(* IEC 61131-3 sources: plcrex/tests/st_to_synchr_models, 21 files *)

(* ---- TC02.st ---- *)
FUNCTION_BLOCK TC02//_functionBlock
  VAR
    x0 : INT;
  END_VAR

  x0 := 0;
END_FUNCTION_BLOCK

(* ---- TC04.st ---- *)
FUNCTION_BLOCK TC04 //_inputs
  VAR_INPUT
    x0 : INT;
    x1 : INT := 6;
  END_VAR
  VAR
    x2 : INT;
  END_VAR

  x2 := x1;
END_FUNCTION_BLOCK

(* ---- TC05.st ---- *)
FUNCTION_BLOCK TC05 //_outputs
  VAR_OUTPUT
    y0 : INT;
    y1 : INT := 6;
  END_VAR
  VAR
    x2 : INT;
  END_VAR

  y0 := x2;
END_FUNCTION_BLOCK

(* ---- TC06.st ---- *)
FUNCTION_BLOCK TC06 //_in_outputs
  VAR_IN_OUT
    y0 : INT;
    y1 : INT;
  END_VAR

  y0 := y1;
END_FUNCTION_BLOCK

(* ---- TC07.st ---- *)
FUNCTION_BLOCK TC07 //_localVariables
  VAR
    x0 : INT;
    x1 : INT := 6;
  END_VAR

  x0 := x1;
END_FUNCTION_BLOCK

(* ---- TC08.st ---- *)
FUNCTION_BLOCK TC08 // _datatypes
  VAR
    x0 : BOOL;
    x1 : BOOL := TRUE;
    x2 : INT;
    x3 : INT := 2;
    x4 : REAL;
    x5 : REAL := 1.23;
    x7 : TIME;
    x8 : TIME := t#5s;
    x9 : ARRAY [1..2] OF BOOL;
    x10 : ARRAY [1..2] OF INT;
    x11 : ARRAY [1..2] OF REAL;
    x12 : ARRAY [1..2] OF TIME;
  END_VAR

  x0 := x1;
  x2 := x3;
  x4 := x5;
  x7 := x8;
  x9[0]:=TRUE;
  x10[0]:=2;
  x11[0]:=1.23;
  x12[0]:=t#2s;
END_FUNCTION_BLOCK

(* ---- TC09.st ---- *)
FUNCTION_BLOCK TC09 //_constants
  VAR
    x0 : BOOL;
    x1 : BOOL := TRUE;
    x2 : BOOL := FALSE;
  END_VAR

  x0 := x1;
  x0 := x2;
END_FUNCTION_BLOCK

(* ---- TC10.st ---- *)
FUNCTION_BLOCK TC10 //Boolean Operators
  VAR
    x0 : BOOL;
    x1 : BOOL := TRUE;
    x2 : BOOL := FALSE;
  END_VAR

  x0 := NOT(x1);
  x0 := x1 AND x2;
  x0 := AND(x1,x2);
  x0 := x1 OR x2;
  x0 := OR(x1,x2);
  x0 := x1 XOR x2;
  x0 := XOR(x1,x2);
END_FUNCTION_BLOCK

(* ---- TC11.st ---- *)
FUNCTION_BLOCK TC11 // _inEquality
  VAR
    x0 : BOOL;
    x1 : BOOL := TRUE;
    x2 : BOOL := FALSE;
  END_VAR

  x0 := x1 = x2;
  x0 := EQ(x1,x2);
  x0 := x1 <> x2;
  x0 := NE(x1,x2);
END_FUNCTION_BLOCK

(* ---- TC12.st ---- *)
FUNCTION_BLOCK TC12 //_numericRelations
  VAR
    x0 : BOOL;
    x1 : INT := 1;
    x2 : INT := 2;
  END_VAR

  x0 := x1 < x2;
  x0 := LT(x1, x2);
  x0 := x1 <= x2;
  x0 := LE(x1, x2);
  x0 := x1 > x2;
  x0 := GT(x1, x2);
  x0 := x1 >= x2;
  x0 := GE(x1, x2);
END_FUNCTION_BLOCK

(* ---- TC13.st ---- *)
FUNCTION_BLOCK TC13 //_arithmeticOperators
  VAR
    x0 : REAL;
    x1 : REAL := 1.0;
    x2 : REAL := 2.0;
    x3 : INT := 1;
    x4 : INT := 2;
    x5 : INT;
  END_VAR

  x0 := x1 + x2;
  x0 := ADD(x1, x2);
  x0 := x1 - x2;
  x0 := SUB(x1, x2);
  x0 := x1 * x2;
  x0 := MUL(x1, x2);
  x0 := x1 / x2;
  x0 := DIV(x1, x2);
  x0 := EXPT(x1, x2);
  x5 := MOD(x3, x4);
END_FUNCTION_BLOCK

(* ---- TC14.st ---- *)
FUNCTION_BLOCK TC14 //_conditional
  VAR
    x0 : BOOL;
    x1 : BOOL := TRUE;
  END_VAR

  IF x1 THEN
    x0:=TRUE;
  ELSE
    x0:= FALSE;
  END_IF;

  x0 := SEL(x1,TRUE,FALSE);
END_FUNCTION_BLOCK

(* ---- TC15.st ---- *)
FUNCTION_BLOCK TC15 //_loop1
  VAR
    x0 : INT := 0;
    x1 : INT := 1;
    y : INT;
    i : INT;
    i0 : INT := 0;
    i1 : INT := 10;
  END_VAR

  i:=i0;
  WHILE i<=i1 DO
    y := x0;
    i := i+1;
  END_WHILE;
  y := x1;
END_FUNCTION_BLOCK

(* ---- TC16.st ---- *)
FUNCTION_BLOCK TC16 // _loop2
  VAR
    x0 : INT := 0;
    x1 : INT := 1;
    y : INT;
    i : INT;
    i0 : INT := 0;
    i1 : INT := 10;
  END_VAR

  i:=i0;
  REPEAT
    y := x0;
    i := i+1;
  UNTIL i>i1
  END_REPEAT;
  y := x1;
END_FUNCTION_BLOCK

(* ---- TC17.st ---- *)
FUNCTION_BLOCK TC17 //_singleAssignment_1
  VAR
    x : INT := 2;
    y : INT;
  END_VAR

  y := x;
END_FUNCTION_BLOCK

(* ---- TC18.st ---- *)
FUNCTION_BLOCK TC18//_singleAssignment_2
  VAR
    x0 : INT := 2;
    x1 : INT := 2;
    y0 : INT;
    y1 : INT;
  END_VAR

  y0 := x0;
  y1 := x1;
END_FUNCTION_BLOCK

(* ---- TC19.st ---- *)
FUNCTION_BLOCK TC19//_multipleAssignment
  VAR
    x0 : INT := 2;
    x1 : INT := 2;
    x2 : INT := 2;
    y1 : INT;
  END_VAR

  y1 := x0;
  y1 := x1;
  y1 := x2;
END_FUNCTION_BLOCK

(* ---- TC20.st ---- *)
FUNCTION_BLOCK TC20//_delayedAssignment
  VAR
    x0 : INT := 2;
    y : INT := 1;
  END_VAR

  y := y + x0;
END_FUNCTION_BLOCK

(* ---- TC21.st ---- *)
FUNCTION_BLOCK TC21
  VAR_OUTPUT
    y : INT;
  END_VAR
  VAR
    x : INT := 1;
    i : INT;
    i0 : INT := 0;
    i1 : INT := 10;
  END_VAR

  i:=i0;
  REPEAT
    y := i;
    i := i+1;
  UNTIL i>i1
  END_REPEAT;
  y := x;
END_FUNCTION_BLOCK

(* ---- TC01.st ---- *)
PROGRAM TC01//_program
  VAR
    x0 : INT;
  END_VAR

  x0 := 0;
END_PROGRAM

(* ---- TC03.st ---- *)
PROGRAM TC03 //_import
  VAR
    fb1 : TC04;
  END_VAR

  fb1(x0 := 2, x1 := 3);
END_PROGRAM
